// TIA Portal V17 export
// export: Created 2026-11-08T05:50:31.9981955Z, ExportSetting WithDefaults, DisplayName Totally Integrated Automation Portal, DisplayVersion V17, DisplayName TIA Portal Openness, DisplayVersion V17, DisplayName TIA Portal Version Control Interface, DisplayVersion V17, DisplayName STEP 7 Professional, DisplayVersion V17, DisplayName STEP 7 Safety, DisplayVersion V17, DisplayName WinCC Professional, DisplayVersion V17
TextList "Estados"  ListRange=Decimal
  TextListEntry   EntryType=SingleValue, Text="REPOSO"
  TextListEntry   EntryType=SingleValue, From=10, To=10, Text="MARCHA"
  TextListEntry   EntryType=SingleValue, From=90, To=90, Text="FALLA"
